FUNCTION_BLOCK T_E_text_Fuse EXTENDS T_E_text_Common
VAR
END_VAR

PROPERTY allFusesOk : KOSTAL_AF2024_Core_Text.ST_E_Text
GET
allFusesOk.Number:= 11;
END_GET
END_PROPERTY

PROPERTY fuse_0_tripped : KOSTAL_AF2024_Core_Text.ST_E_Text
GET
fuse_0_tripped.Number:= 10;
END_GET
END_PROPERTY

PROPERTY name : KOSTAL_AF2024_Core_Text.ST_E_Text
GET
name.Number:= 2;
END_GET
END_PROPERTY

END_FUNCTION_BLOCK

(* stored: Version 1.1.0.1, ProductVersion 3.1.4024.12
   POU T_E_text_Fuse: Id {c8a49c64-d262-4349-b63a-ac422e401bc8}, SpecialFunc None
   Property allFusesOk: Id {21bb1c91-a78a-4577-861d-a4c0a08af0a6}
   Get Get: Id {deacaa57-d416-4eaf-be50-8022c70fb033}
   Property fuse_0_tripped: Id {8f62ed67-06e6-4e19-9b45-4e9d99de17f8}
   Get Get: Id {2201fcf2-6757-4bf2-ae80-c395954698b3}
   Property name: Id {81c95c70-60ef-42bb-bfd9-abe58fa5b682}
   Get Get: Id {5811258e-0bb4-44b8-9423-124d411851b3} *)
